(* IEC 61131-3 sources: JingjiangArm/moonboxpro_arm_8.4/Application/Application/数据类型/枚举, 4 files *)

(* ---- ENUM_LogicRunSteps.st ---- *)
(*@CES
Name=ENUM_LogicRunSteps
Type=Gvl
TypeGuid=2db5746d-d284-4425-9f7f-2663a34b0ebc
Guid=7d453960-5c1c-45de-90db-0b154bc5d5ec
HasDeclaration=True
HasImplementation=False
*)
{DECLARATION}
TYPE ENUM_LogicRunSteps :
(
	RUNSTEP_STARTUP					,(*初始化内容*)
	RUNSTEP_RdRingNetStationDetails	,(* 读取驱动器所有的相关信息 *)
	RUNSTEP_LoadSysParam			,(* 装载系统参数 *)
	RUNSTEP_LoadSysCfg				,(* 加载系统配置/2021.11.29.181715/hdp *)
	RUNSTEP_UpdateSysCfg			,(* 更新系统配置/2021.11.29.181715/hdp *)
	RUNSTEP_LoadCfg_Motor			,(* 过渡状态 *)
	RUNSTEP_NormalWork				,(* 正常工作状态 *)
(*deprecated@2021.12.21.163944/hdp
	RUNSTEP_Enter_Cfg_Wizard		,(* 进入系统配置的向导页/2021.11.29.174122/hdp *)
*)
(*deprecated@2021.12.21.161925/hdp
	RUNSTEP_Enter_Param_Wizard		,(* 进入系统参数的向导页/2021.11.29.174122/hdp *)
*)
	RUNSTEP_SETMODAL				,(*2024.10.25.083548设置模态*)
	RUNSTEP_RESERVED				 (* 保留 *)
);
END_TYPE

{IMPLEMENTATION}

(* ---- ENUM_MarkArrangeType.st ---- *)
(*@CES
Name=ENUM_MarkArrangeType
Type=Gvl
TypeGuid=2db5746d-d284-4425-9f7f-2663a34b0ebc
Guid=1b9c9704-f7e9-4499-af37-1e699b1dbe55
HasDeclaration=True
HasImplementation=False
*)
{DECLARATION}
TYPE ENUM_MarkArrangeType :
(
	MARK_ARRANGE_VFOR		:= 1, (* 纵顺 *)
	MARK_ARRANGE_VREV		:= 2, (* 纵逆 *)
	MARK_ARRANGE_HFOR		:= 3, (* 横顺 *)
	MARK_ARRANGE_HREV		:= 4, (* 横逆 *)
	MARK_ARRANGE_OMK		:= 5  (* 单标记 *)
);
END_TYPE

{IMPLEMENTATION}

(* ---- ENUM_MarkType.st ---- *)
(*@CES
Name=ENUM_MarkType
Type=Gvl
TypeGuid=2db5746d-d284-4425-9f7f-2663a34b0ebc
Guid=321db1e3-f3d5-4ccd-ba69-c64547f2641d
HasDeclaration=True
HasImplementation=False
*)
{DECLARATION}
TYPE ENUM_MarkType :
(
	MARK_TYPE_LINE			:= 1, (* Line Mark *)
	MARK_TYPE_TRAPE_VFLP	:= 2, (* Vert Forward Left Positive *)
	MARK_TYPE_TRAPE_VFLN	:= 3, (* Vert Forward Left Negitive *)
	MARK_TYPE_TRAPE_VBLP	:= 4, (* Vert Backward Left Positive *)
	MARK_TPYE_TRAPE_VBLN	:= 5, (* Vert Backward Left Negitive *)
	MARK_TYPE_TRIANGLE_R	:= 6, (* 2018.8.28.135823\三角标-定点在右边 *)
	MARK_TYPE_TRIANGLE_L	:= 7  (* 2018.8.28.135828\三角标-定点在左边 *)
);
END_TYPE

{IMPLEMENTATION}

(* ---- ENUMS_STEP_RDRINGNET.st ---- *)
(*@CES
Name=ENUMS_STEP_RDRINGNET
Type=Gvl
TypeGuid=2db5746d-d284-4425-9f7f-2663a34b0ebc
Guid=ae3e14f3-c75e-4491-bf67-9f081b73171a
HasDeclaration=True
HasImplementation=False
*)
{DECLARATION}
TYPE ENUMS_STEP_RDRINGNET :
(
	CASE_STANDBY				:= -1,(* 默认就绪状态 *)
	CASE_GET_RINGNET_INF		:= 1,(* 读取等环网网络信息 *)
	CASE_GET_DRV_TYPE			:= 2,(* 读取驱动器的型号 *)
	CASE_GET_DRV_PWR_LEVEL		:= 3,(* 读取驱动器的功率等级 *)
	CASE_GET_DRV_FW_VERSION		:= 4,(* 读取驱动器的固件版本 *)
	CASE_GET_DRV_PARAM_NRS		:= 5,(* 读取电机的额定转速 *)
	CASE_GET_DRV_PARAM_NOS		:= 6,(* 读取电机的过速转速 *)
	CASE_GET_DRV_PARAM_IMAX		:= 7,(* 读取电机的最大电流 *)
	CASE_GET_DRV_PARAM_POSOFST	:= 8,(* 读取位置偏移 *)
	CASE_GEN_SUMMARY_OF_STATION	:= 9,(* 生成有关站号的摘要信息 *)
	CASE_GET_DRV_PARAM_TORQUE	:= 10(* 读取扭矩系数 *)
);
END_TYPE

{IMPLEMENTATION}
